{attribute 'qualified_only'}
VAR_GLOBAL CONSTANT
	MAX_VALVES		: INT := 8;
	DEFAULT_TIMEOUT	: TIME := T#5S;
END_VAR

(* stored: Version 1.1.0.1
   GVL GVL_DemoLib: Id {d61f31a9-324a-4c9c-add8-0db271036033} *)
